Fanuc KAREL source: KT00495.KL

PROGRAM KT00495
%NOLOCKGROUP
VAR
  P1: XYZWPR
  P2: POSITION
  OUT: XYZWPR
BEGIN
  P1.X = 1.0
  OUT = P1 : P2
END KT00495
